// TIA Portal V19 export
FUNCTION_BLOCK "ALL_VALVES"   // FB1, FBD
{ S7_Optimized_Access := 'TRUE' }
// stored: MemoryReserve 100, SetENOAutomatically false
   VAR
      XV01 { S7_SetPoint := 'True'} : "valve";
      XV02 { S7_SetPoint := 'True'} : "valve";
      XV03 { S7_SetPoint := 'True'} : "valve";
      XV04 { S7_SetPoint := 'True'} : "valve";
      XV05 { S7_SetPoint := 'True'} : "valve";
      XV06 { S7_SetPoint := 'True'} : "valve";
      XV07 { S7_SetPoint := 'True'} : "valve";
      XV08 { S7_SetPoint := 'True'} : "valve";
   END_VAR
BEGIN

REGION Network 1
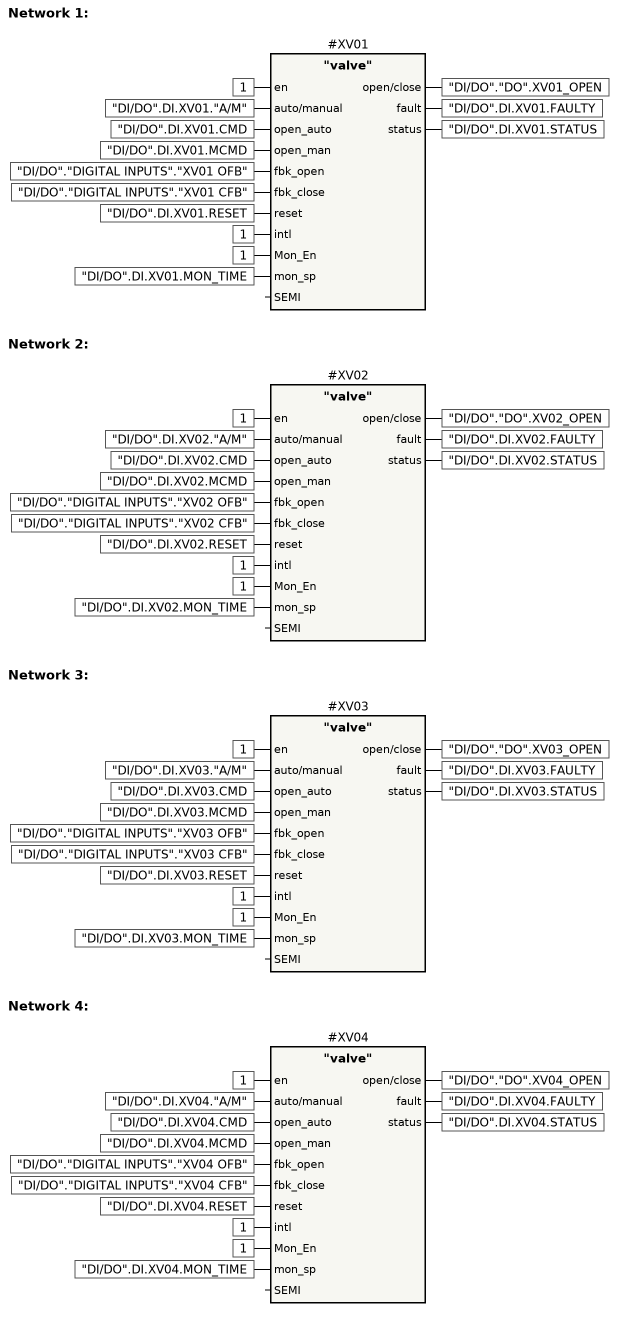
   IF 1 THEN
       #XV01("auto/manual" := "DI/DO".DI.XV01."A/M",   // "valve"
             open_auto := "DI/DO".DI.XV01.CMD,
             open_man := "DI/DO".DI.XV01.MCMD,
             fbk_open := "DI/DO"."DIGITAL INPUTS"."XV01 OFB",
             fbk_close := "DI/DO"."DIGITAL INPUTS"."XV01 CFB",
             reset := "DI/DO".DI.XV01.RESET,
             intl := 1,
             Mon_En := 1,
             mon_sp := "DI/DO".DI.XV01.MON_TIME,
             "open/close" => "DI/DO"."DO".XV01_OPEN,
             fault => "DI/DO".DI.XV01.FAULTY,
             status => "DI/DO".DI.XV01.STATUS);
   END_IF;
END_REGION

REGION Network 2
   IF 1 THEN
       #XV02("auto/manual" := "DI/DO".DI.XV02."A/M",   // "valve"
             open_auto := "DI/DO".DI.XV02.CMD,
             open_man := "DI/DO".DI.XV02.MCMD,
             fbk_open := "DI/DO"."DIGITAL INPUTS"."XV02 OFB",
             fbk_close := "DI/DO"."DIGITAL INPUTS"."XV02 CFB",
             reset := "DI/DO".DI.XV02.RESET,
             intl := 1,
             Mon_En := 1,
             mon_sp := "DI/DO".DI.XV02.MON_TIME,
             "open/close" => "DI/DO"."DO".XV02_OPEN,
             fault => "DI/DO".DI.XV02.FAULTY,
             status => "DI/DO".DI.XV02.STATUS);
   END_IF;
END_REGION

REGION Network 3
   IF 1 THEN
       #XV03("auto/manual" := "DI/DO".DI.XV03."A/M",   // "valve"
             open_auto := "DI/DO".DI.XV03.CMD,
             open_man := "DI/DO".DI.XV03.MCMD,
             fbk_open := "DI/DO"."DIGITAL INPUTS"."XV03 OFB",
             fbk_close := "DI/DO"."DIGITAL INPUTS"."XV03 CFB",
             reset := "DI/DO".DI.XV03.RESET,
             intl := 1,
             Mon_En := 1,
             mon_sp := "DI/DO".DI.XV03.MON_TIME,
             "open/close" => "DI/DO"."DO".XV03_OPEN,
             fault => "DI/DO".DI.XV03.FAULTY,
             status => "DI/DO".DI.XV03.STATUS);
   END_IF;
END_REGION

REGION Network 4
   IF 1 THEN
       #XV04("auto/manual" := "DI/DO".DI.XV04."A/M",   // "valve"
             open_auto := "DI/DO".DI.XV04.CMD,
             open_man := "DI/DO".DI.XV04.MCMD,
             fbk_open := "DI/DO"."DIGITAL INPUTS"."XV04 OFB",
             fbk_close := "DI/DO"."DIGITAL INPUTS"."XV04 CFB",
             reset := "DI/DO".DI.XV04.RESET,
             intl := 1,
             Mon_En := 1,
             mon_sp := "DI/DO".DI.XV04.MON_TIME,
             "open/close" => "DI/DO"."DO".XV04_OPEN,
             fault => "DI/DO".DI.XV04.FAULTY,
             status => "DI/DO".DI.XV04.STATUS);
   END_IF;
END_REGION

REGION Network 5
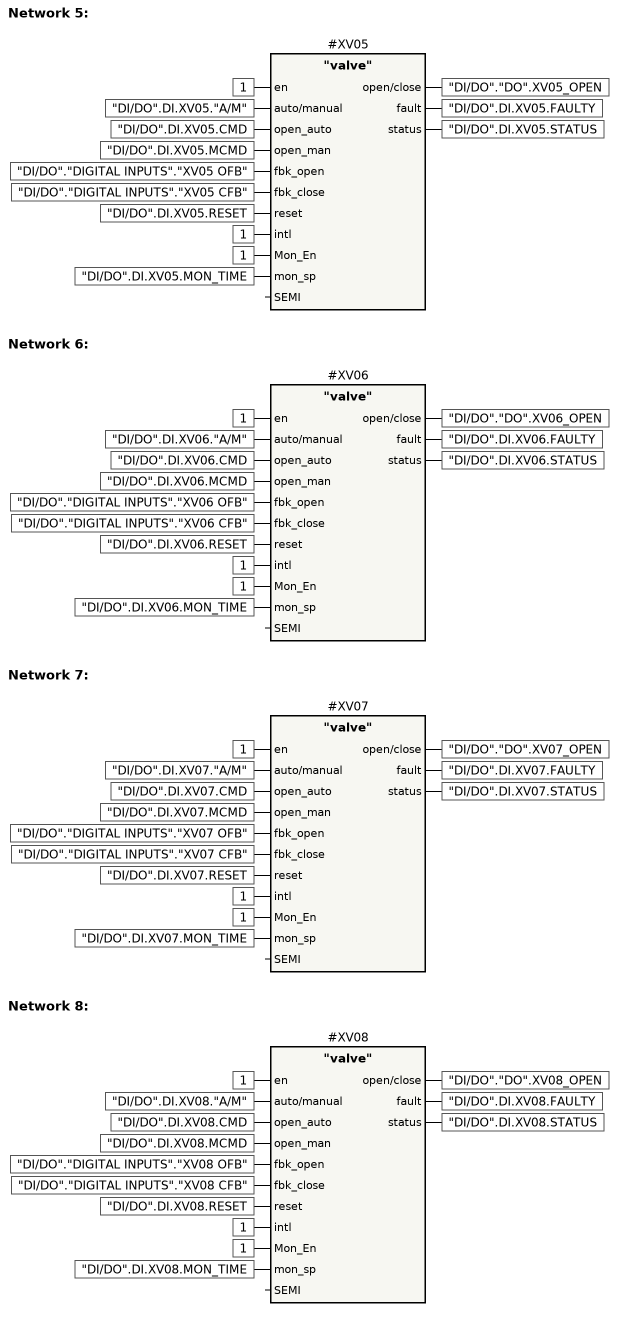
   IF 1 THEN
       #XV05("auto/manual" := "DI/DO".DI.XV05."A/M",   // "valve"
             open_auto := "DI/DO".DI.XV05.CMD,
             open_man := "DI/DO".DI.XV05.MCMD,
             fbk_open := "DI/DO"."DIGITAL INPUTS"."XV05 OFB",
             fbk_close := "DI/DO"."DIGITAL INPUTS"."XV05 CFB",
             reset := "DI/DO".DI.XV05.RESET,
             intl := 1,
             Mon_En := 1,
             mon_sp := "DI/DO".DI.XV05.MON_TIME,
             "open/close" => "DI/DO"."DO".XV05_OPEN,
             fault => "DI/DO".DI.XV05.FAULTY,
             status => "DI/DO".DI.XV05.STATUS);
   END_IF;
END_REGION

REGION Network 6
   IF 1 THEN
       #XV06("auto/manual" := "DI/DO".DI.XV06."A/M",   // "valve"
             open_auto := "DI/DO".DI.XV06.CMD,
             open_man := "DI/DO".DI.XV06.MCMD,
             fbk_open := "DI/DO"."DIGITAL INPUTS"."XV06 OFB",
             fbk_close := "DI/DO"."DIGITAL INPUTS"."XV06 CFB",
             reset := "DI/DO".DI.XV06.RESET,
             intl := 1,
             Mon_En := 1,
             mon_sp := "DI/DO".DI.XV06.MON_TIME,
             "open/close" => "DI/DO"."DO".XV06_OPEN,
             fault => "DI/DO".DI.XV06.FAULTY,
             status => "DI/DO".DI.XV06.STATUS);
   END_IF;
END_REGION

REGION Network 7
   IF 1 THEN
       #XV07("auto/manual" := "DI/DO".DI.XV07."A/M",   // "valve"
             open_auto := "DI/DO".DI.XV07.CMD,
             open_man := "DI/DO".DI.XV07.MCMD,
             fbk_open := "DI/DO"."DIGITAL INPUTS"."XV07 OFB",
             fbk_close := "DI/DO"."DIGITAL INPUTS"."XV07 CFB",
             reset := "DI/DO".DI.XV07.RESET,
             intl := 1,
             Mon_En := 1,
             mon_sp := "DI/DO".DI.XV07.MON_TIME,
             "open/close" => "DI/DO"."DO".XV07_OPEN,
             fault => "DI/DO".DI.XV07.FAULTY,
             status => "DI/DO".DI.XV07.STATUS);
   END_IF;
END_REGION

REGION Network 8
   IF 1 THEN
       #XV08("auto/manual" := "DI/DO".DI.XV08."A/M",   // "valve"
             open_auto := "DI/DO".DI.XV08.CMD,
             open_man := "DI/DO".DI.XV08.MCMD,
             fbk_open := "DI/DO"."DIGITAL INPUTS"."XV08 OFB",
             fbk_close := "DI/DO"."DIGITAL INPUTS"."XV08 CFB",
             reset := "DI/DO".DI.XV08.RESET,
             intl := 1,
             Mon_En := 1,
             mon_sp := "DI/DO".DI.XV08.MON_TIME,
             "open/close" => "DI/DO"."DO".XV08_OPEN,
             fault => "DI/DO".DI.XV08.FAULTY,
             status => "DI/DO".DI.XV08.STATUS);
   END_IF;
END_REGION
END_FUNCTION_BLOCK
